(* IEC 61131-3 sources: volt/packages/volt-lsp-iec/test-corpus/bakon-nano/Device/Plc Logic/Application/Library Manager/StringUtils, 84 files *)

(* ---- CHARBUFFERPTR.dut ---- *)
TYPE CHARBUFFERPTR : POINTER TO BYTE;
END_TYPE

(* ---- DATETIMEPLACEHOLDEROCCURRENCE.dut ---- *)
TYPE DATETIMEPLACEHOLDEROCCURRENCE :
STRUCT
	M_EPLACEHOLDER : EDateTimePlaceholder;
	M_IOFFSET : INT;
	M_ILENGTH : INT;
END_STRUCT
END_TYPE

(* ---- EDATETIMEPLACEHOLDER.dut ---- *)
TYPE EDATETIMEPLACEHOLDER :
(
	PLH_IS_VALID := 0,
	DFMT_5_DIGIT_DAY := 40,
	DFMT_4_DIGIT_DAY := 41,
	DFMT_3_DIGIT_DAY := 42,
	DFMT_2_DIGIT_DAY := 43,
	DFMT_1_DIGIT_DAY := 44,
	DFMT_3_DIGIT_DAYOFYEAR := 45,
	DFMT_4_DIGIT_MONTH := 46,
	DFMT_3_DIGIT_MONTH := 47,
	DFMT_2_DIGIT_MONTH := 48,
	DFMT_1_DIGIT_MONTH := 49,
	DFMT_4_DIGIT_YEAR := 50,
	DFMT_2_DIGIT_YEAR := 51,
	DFMT_1_DIGIT_YEAR := 52,
	TFMT_2_DIGIT_HOUR_24_HOUR_CLOCK := 60,
	TFMT_1_DIGIT_HOUR_24_HOUR_CLOCK := 61,
	TFMT_2_DIGIT_HOUR_12_HOUR_CLOCK := 62,
	TFMT_1_DIGIT_HOUR_12_HOUR_CLOCK := 63,
	TFMT_3_DIGIT_MILLISECOND := 64,
	TFMT_3_DIGIT_MICROSECOND := 65,
	TFMT_3_DIGIT_NANOSECOND := 66,
	TFMT_2_DIGIT_MINUTE := 67,
	TFMT_1_DIGIT_MINUTE := 68,
	TFMT_2_DIGIT_SECOND := 69,
	TFMT_1_DIGIT_SECOND := 70,
	TFMT_AM_PM_DESIGNATOR := 71,
	TFMT_1_DIGIT_AM_PM_DESIGNATOR := 72,
	TFMT_1_DIGIT_ZONE_DESIGNATOR := 73,
	PLH_NOT_USED := 255
);
END_TYPE

(* ---- EPLACEHOLDERANALYZATIONSTATE.dut ---- *)
TYPE EPLACEHOLDERANALYZATIONSTATE :
(
	NOTAVAILABLE := 16#0,
	TOOMANYPLACEHOLDERS := 16#1,
	DONE := 16#10
);
END_TYPE

(* ---- PLACEHOLDERDESCRIPTION.dut ---- *)
TYPE PLACEHOLDERDESCRIPTION :
STRUCT
	M_EPLACEHOLDER : EDateTimePlaceholder;
	M_PCBSPLACEHOLDER : POINTER TO CharBufferString;
	M_XCONSIDERPLACEHOLDER : BOOL := TRUE;
	M_PRELATEDPLACEHOLDERISSUBSTRINGOF : POINTER TO PlaceholderDescription;
	M_PRELATEDPLACEHOLDERHASSUBSTRING : POINTER TO PlaceholderDescription;
END_STRUCT
END_TYPE

(* ---- CONSTANTS.gvl ---- *)
VAR_GLOBAL
	NULL : POINTER TO BYTE := 0;
END_VAR

(* ---- GVL_UTF8.gvl ---- *)
VAR_GLOBAL
	TRAILINGBYTESFORUTF8 : ARRAY [0..255] OF BYTE := [0, 0, 0, 0, 0, 0, 0, 0, 0, 0, 0, 0, 0, 0, 0, 0, 0, 0, 0, 0, 0, 0, 0, 0, 0, 0, 0, 0, 0, 0, 0, 0, 0, 0, 0, 0, 0, 0, 0, 0, 0, 0, 0, 0, 0, 0, 0, 0, 0, 0, 0, 0, 0, 0, 0, 0, 0, 0, 0, 0, 0, 0, 0, 0, 0, 0, 0, 0, 0, 0, 0, 0, 0, 0, 0, 0, 0, 0, 0, 0, 0, 0, 0, 0, 0, 0, 0, 0, 0, 0, 0, 0, 0, 0, 0, 0, 0, 0, 0, 0, 0, 0, 0, 0, 0, 0, 0, 0, 0, 0, 0, 0, 0, 0, 0, 0, 0, 0, 0, 0, 0, 0, 0, 0, 0, 0, 0, 0, 0, 0, 0, 0, 0, 0, 0, 0, 0, 0, 0, 0, 0, 0, 0, 0, 0, 0, 0, 0, 0, 0, 0, 0, 0, 0, 0, 0, 0, 0, 0, 0, 0, 0, 0, 0, 0, 0, 0, 0, 0, 0, 0, 0, 0, 0, 0, 0, 0, 0, 0, 0, 0, 0, 0, 0, 0, 0, 0, 0, 0, 0, 0, 0, 1, 1, 1, 1, 1, 1, 1, 1, 1, 1, 1, 1, 1, 1, 1, 1, 1, 1, 1, 1, 1, 1, 1, 1, 1, 1, 1, 1, 1, 1, 1, 1, 2, 2, 2, 2, 2, 2, 2, 2, 2, 2, 2, 2, 2, 2, 2, 2, 3, 3, 3, 3, 3, 3, 3, 3, 4, 4, 4, 4, 5, 5, 5, 5];
	FIRSTBYTEMARK : ARRAY [0..6] OF BYTE := [16#0, 16#0, 16#C0, 16#E0, 16#F0, 16#F8, 16#FC];
	OFFSETSFROMUTF8 : ARRAY [0..5] OF DWORD := [16#0, 16#3080, 16#E2080, 16#3C82080, 16#FA082080, 16#82082080];
	HALFSHIFT : INT := 10;
	HALFBASE : DWORD := 16#10000;
	HALFMASK : DWORD := 16#3FF;
	UNI_REPLACEMENT_CHAR : DWORD := 16#FFFD;
	UNI_MAX_BMP : DWORD := 16#FFFF;
	UNI_MAX_UTF16 : DWORD := 16#10FFFF;
	UNI_MAX_UTF32 : DWORD := 16#7FFFFFFF;
	UNI_MAX_LEGAL_UTF32 : DWORD := 16#10FFFF;
	BYTEMASK : DWORD := 16#BF;
	BYTEMARK : DWORD := 16#80;
	UNI_SUR_HIGH_START : DWORD := 16#D800;
	UNI_SUR_HIGH_END : DWORD := 16#DBFF;
	UNI_SUR_LOW_START : DWORD := 16#DC00;
	UNI_SUR_LOW_END : DWORD := 16#DFFF;
	ERR_SOURCE_EXHAUSTED : UDINT := 16#40A0;
	ERR_TARGET_EXHAUSTED : UDINT := 16#40A1;
	ERR_SOURCE_ILLEGAL : UDINT := 16#40A2;
END_VAR

(* ---- PLACEHOLDERCONSTANTS.gvl ---- *)
VAR_GLOBAL
	DFMT_FIRST_PLACEHOLDER : EDateTimePlaceholder := EDateTimePlaceholder.DFMT_5_DIGIT_DAY;
	DFMT_LAST_PLACEHOLDER : EDateTimePlaceholder := EDateTimePlaceholder.DFMT_1_DIGIT_YEAR;
	TFMT_FIRST_PLACEHOLDER : EDateTimePlaceholder := EDateTimePlaceholder.TFMT_2_DIGIT_HOUR_24_HOUR_CLOCK;
	TFMT_LAST_PLACEHOLDER : EDateTimePlaceholder := EDateTimePlaceholder.TFMT_1_DIGIT_ZONE_DESIGNATOR;
END_VAR

(* ---- STRINGUTILSVERSIONCONSTANTS.gvl ---- *)
VAR_GLOBAL
	_STRINGUTILS_VERSION_LARGEROREQUAL_3_5_3_40_ : INT := 0;
END_VAR

(* ---- ICHARBUFFERSTRING.itf ---- *)
INTERFACE ICHARBUFFERSTRING
END_INTERFACE

METHOD ASWSTRING : CharBufferPtr
END_METHOD

METHOD COPY : DINT
VAR_INPUT
	CBSSOURCE : REFERENCE TO CharBufferString;
END_VAR
END_METHOD

METHOD FROMSTRING : BOOL
VAR_INPUT
	STSTRING : STRING(255);
END_VAR
END_METHOD

METHOD INITCONVERTED : BOOL
VAR_INPUT
	PBUFFER : POINTER TO BYTE;
	UIBUFFERSIZE : UINT;
END_VAR
END_METHOD

(* ---- ILOCALIZEDDATETIMENAMES.itf ---- *)
INTERFACE ILOCALIZEDDATETIMENAMES
END_INTERFACE

METHOD GETDAYLONG : CharBufferPtr
VAR_INPUT
	UIDAYOFWEEK : UINT;
END_VAR
END_METHOD

METHOD GETDAYSHORT : CharBufferPtr
VAR_INPUT
	UIDAYOFWEEK : UINT;
END_VAR
END_METHOD

METHOD GETMONTHLONG : CharBufferPtr
VAR_INPUT
	UIMONTH : UINT;
END_VAR
END_METHOD

METHOD GETMONTHSHORT : CharBufferPtr
VAR_INPUT
	UIMONTH : UINT;
END_VAR
END_METHOD

(* ---- _PRINTF.pou ---- *)
FUNCTION _PRINTF : BOOL
VAR_INPUT
	CBPRESULT : CharBufferPtr;
	UIRESULTCAPACITY : UINT;
	STRINGTYPE : __SYSTEM.TYPE_CLASS;
	CBPFORMAT : CharBufferPtr;
	PVALUE : POINTER TO BYTE;
	TYPECLASS : __SYSTEM.TYPE_CLASS;
END_VAR
END_FUNCTION

(* ---- ANALYZEPLACEHOLDERS.pou ---- *)
FUNCTION ANALYZEPLACEHOLDERS : EPlaceholderAnalyzationState
VAR_INPUT
	RCBSMESSAGE : REFERENCE TO CharBufferString;
	PAPLACEHOLDERS : POINTER TO ARRAY [0..0] OF PlaceholderDescription;
	ICOUNTPLACEHOLDERTOCHECK : INT;
	PAPLACEHOLDEROCCURRENCE : POINTER TO ARRAY [0..0] OF DateTimePlaceholderOccurrence;
	SIMAXCOUNTPLACEHOLDERS : SINT;
END_VAR
VAR_OUTPUT
	SICOUNTPLACEHOLDERS : SINT;
END_VAR
END_FUNCTION

(* ---- ANALYZEPLACEHOLDERSDATETIME.pou ---- *)
FUNCTION ANALYZEPLACEHOLDERSDATETIME : EPlaceholderAnalyzationState
VAR_INPUT
	RCBSMESSAGE : REFERENCE TO CharBufferString;
	PAPLACEHOLDERS : POINTER TO ARRAY [0..0] OF PlaceholderDescription;
	ICOUNTPLACEHOLDERTOCHECK : INT;
	PAPLACEHOLDEROCCURRENCE : POINTER TO ARRAY [0..0] OF DateTimePlaceholderOccurrence;
	SIMAXCOUNTPLACEHOLDERS : SINT;
END_VAR
VAR_OUTPUT
	SICOUNTPLACEHOLDERS : SINT;
END_VAR
END_FUNCTION

(* ---- CHARACTERATEQUALS.pou ---- *)
FUNCTION CHARACTERATEQUALS : BOOL
VAR_INPUT
	CBSSOURCE : REFERENCE TO CharBufferString;
	IPOSITION : INT;
	STCHAR : STRING(1);
END_VAR
END_FUNCTION

(* ---- CHARTOUPPER.pou ---- *)
FUNCTION CHARTOUPPER : BYTE
VAR_INPUT
	BYCHAR : BYTE;
END_VAR
END_FUNCTION

(* ---- CONVERTUTF16TOUTF8.pou ---- *)
FUNCTION CONVERTUTF16TOUTF8 : UDINT
VAR_INPUT
	SOURCESTART : POINTER TO WORD;
	TARGETSTART : POINTER TO BYTE;
	DWTARGETBUFFERSIZE : DWORD;
	BSTRICTCONVERSION : BOOL;
END_VAR
END_FUNCTION

(* ---- CONVERTUTF8TOUTF16.pou ---- *)
FUNCTION CONVERTUTF8TOUTF16 : UDINT
VAR_INPUT
	SOURCESTART : POINTER TO BYTE;
	TARGETSTART : POINTER TO WORD;
	DWTARGETBUFFERSIZE : DWORD;
	BSTRICTCONVERSION : BOOL;
END_VAR
END_FUNCTION

(* ---- HELPISSAMEIGNORECASE.pou ---- *)
FUNCTION HELPISSAMEIGNORECASE : BOOL
VAR_INPUT
	BY1 : BYTE;
	BY2 : BYTE;
END_VAR
END_FUNCTION

(* ---- HELPSTRCMPENDA.pou ---- *)
FUNCTION HELPSTRCMPENDA : BOOL
VAR_INPUT
	PCOMPLETETEXT : CharBufferPtr;
	PSUBTEXT : CharBufferPtr;
	XIGNORECASE : BOOL;
END_VAR
END_FUNCTION

(* ---- HELPSTRCMPSTARTA.pou ---- *)
FUNCTION HELPSTRCMPSTARTA : BOOL
VAR_INPUT
	PCOMPLETETEXT : CharBufferPtr;
	PSUBTEXT : CharBufferPtr;
	XIGNORECASE : BOOL;
END_VAR
END_FUNCTION

(* ---- HELPTRIM.pou ---- *)
FUNCTION HELPTRIM : POINTER TO BYTE
VAR_INPUT
	PTEXT : CharBufferPtr;
	XTRIMLEFT : BOOL;
END_VAR
END_FUNCTION

(* ---- HELPTRIMW.pou ---- *)
FUNCTION HELPTRIMW : POINTER TO WORD
VAR_INPUT
	PTEXT : CharBufferPtr;
	XTRIMLEFT : BOOL;
END_VAR
END_FUNCTION

(* ---- ISLEGALUTF8.pou ---- *)
FUNCTION ISLEGALUTF8 : BOOL
VAR_INPUT
	SOURCE : POINTER TO BYTE;
	LENGTH : INT;
END_VAR
END_FUNCTION

(* ---- ISSPACECHARACTER.pou ---- *)
FUNCTION ISSPACECHARACTER : BOOL
VAR_INPUT
	WCHARACTER : WORD;
END_VAR
END_FUNCTION

(* ---- PRINTF.pou ---- *)
FUNCTION PRINTF
VAR_INPUT
	CBSRESULT : REFERENCE TO CharBufferString;
	CBSFORMAT : REFERENCE TO CharBufferString;
	PVALUE : POINTER TO BYTE;
	TYPECLASS : __SYSTEM.TYPE_CLASS;
END_VAR
END_FUNCTION

(* ---- STRATOW.pou ---- *)
FUNCTION STRATOW
VAR_INPUT
	PBYTARGETW : POINTER TO BYTE;
	IBUFFERSIZE : DINT;
	PBYSOURCEA : POINTER TO BYTE;
END_VAR
END_FUNCTION

(* ---- STRCASECMPA.pou ---- *)
FUNCTION STRCASECMPA : INT
VAR_INPUT
	PBYTE1 : POINTER TO BYTE;
	PBYTE2 : POINTER TO BYTE;
END_VAR
END_FUNCTION

(* ---- STRCASECMPENDA.pou ---- *)
FUNCTION STRCASECMPENDA : INT
VAR_INPUT
	PSTRING : CharBufferPtr;
	PSUFFIX : CharBufferPtr;
END_VAR
END_FUNCTION

(* ---- STRCASECMPSTARTA.pou ---- *)
FUNCTION STRCASECMPSTARTA : INT
VAR_INPUT
	PSTRING : CharBufferPtr;
	PPREFIX : CharBufferPtr;
END_VAR
END_FUNCTION

(* ---- STRCASECMPW.pou ---- *)
FUNCTION STRCASECMPW : INT
VAR_INPUT
	PWD1 : POINTER TO WORD;
	PWD2 : POINTER TO WORD;
END_VAR
END_FUNCTION

(* ---- STRCASEFINDA.pou ---- *)
FUNCTION STRCASEFINDA : INT
VAR_INPUT
	PST1 : POINTER TO STRING(255);
	PST2 : POINTER TO STRING(255);
	UISEARCHSTART : UINT;
END_VAR
END_FUNCTION

(* ---- STRCASEFINDW.pou ---- *)
FUNCTION STRCASEFINDW : INT
VAR_INPUT
	PST1 : POINTER TO WSTRING(255);
	PST2 : POINTER TO WSTRING(255);
	UISEARCHSTART : UINT;
END_VAR
END_FUNCTION

(* ---- STRCMP.pou ---- *)
FUNCTION STRCMP : DINT
VAR_INPUT
	CBSSTRING1 : REFERENCE TO CharBufferString;
	CBSSTRING2 : REFERENCE TO CharBufferString;
END_VAR
END_FUNCTION

(* ---- STRCMPA.pou ---- *)
FUNCTION STRCMPA : INT
VAR_INPUT
	PBY1 : POINTER TO BYTE;
	PBY2 : POINTER TO BYTE;
END_VAR
END_FUNCTION

(* ---- STRCMPENDA.pou ---- *)
FUNCTION STRCMPENDA : INT
VAR_INPUT
	PSTRING : CharBufferPtr;
	PSUFFIX : CharBufferPtr;
END_VAR
END_FUNCTION

(* ---- STRCMPSTARTA.pou ---- *)
FUNCTION STRCMPSTARTA : INT
VAR_INPUT
	PSTRING : CharBufferPtr;
	PPREFIX : CharBufferPtr;
END_VAR
END_FUNCTION

(* ---- STRCMPW.pou ---- *)
FUNCTION STRCMPW : INT
VAR_INPUT
	PWD1 : POINTER TO WORD;
	PWD2 : POINTER TO WORD;
END_VAR
END_FUNCTION

(* ---- STRCONCATA.pou ---- *)
FUNCTION STRCONCATA : BOOL
VAR_INPUT
	PSTFROM : CharBufferPtr;
	PSTTO : CharBufferPtr;
	IBUFFERSIZE : INT;
END_VAR
END_FUNCTION

(* ---- STRCONCATW.pou ---- *)
FUNCTION STRCONCATW : BOOL
VAR_INPUT
	PSTFROM : CharBufferPtr;
	PSTTO : CharBufferPtr;
	IBUFFERSIZE : INT;
END_VAR
END_FUNCTION

(* ---- STRCPY.pou ---- *)
FUNCTION STRCPY : DINT
VAR_INPUT
	CBSTARGET : REFERENCE TO CharBufferString;
	CBSSOURCE : REFERENCE TO CharBufferString;
END_VAR
END_FUNCTION

(* ---- STRCPYA.pou ---- *)
FUNCTION STRCPYA : DINT
VAR_INPUT
	PBUFFER : CharBufferPtr;
	IBUFFERSIZE : DINT;
	PSTR : CharBufferPtr;
END_VAR
END_FUNCTION

(* ---- STRCPYFROM.pou ---- *)
FUNCTION STRCPYFROM : DINT
VAR_INPUT
	RCBSTARGET : REFERENCE TO CharBufferString;
	RCBSSOURCE : REFERENCE TO CharBufferString;
	DISOURCEOFFSET : DINT;
	DITARGETOFFSET : DINT;
	DICOUNTCHARACTERS : DINT;
END_VAR
END_FUNCTION

(* ---- STRCPYW.pou ---- *)
FUNCTION STRCPYW : DINT
VAR_INPUT
	PBUFFER : CharBufferPtr;
	IBUFFERSIZE : DINT;
	PSTR : CharBufferPtr;
END_VAR
END_FUNCTION

(* ---- STRDELETE.pou ---- *)
FUNCTION STRDELETE
VAR_INPUT
	CBSSOURCE : REFERENCE TO CharBufferString;
	ILENGTH : INT;
	IPOSITION : INT;
END_VAR
END_FUNCTION

(* ---- STRDELETEA.pou ---- *)
FUNCTION STRDELETEA
VAR_INPUT
	PBY : POINTER TO BYTE;
	ILENGTH : INT;
	IPOSITION : INT;
END_VAR
END_FUNCTION

(* ---- STRDELETEW.pou ---- *)
FUNCTION STRDELETEW
VAR_INPUT
	PWD : POINTER TO WORD;
	ILENGTH : INT;
	IPOSITION : INT;
END_VAR
END_FUNCTION

(* ---- STRFIND.pou ---- *)
FUNCTION STRFIND : INT
VAR_INPUT
	CBSSOURCE : REFERENCE TO CharBufferString;
	CBSTOSEARCHFOR : REFERENCE TO CharBufferString;
END_VAR
END_FUNCTION

(* ---- STRFINDA.pou ---- *)
FUNCTION STRFINDA : INT
VAR_INPUT
	PST1 : POINTER TO STRING(255);
	PST2 : POINTER TO STRING(255);
	UISEARCHSTART : UINT;
END_VAR
END_FUNCTION

(* ---- STRFINDFROM.pou ---- *)
FUNCTION STRFINDFROM : INT
VAR_INPUT
	CBSSOURCE : REFERENCE TO CharBufferString;
	CBSTOSEARCHFOR : REFERENCE TO CharBufferString;
	ISEARCHSTART : UINT;
END_VAR
END_FUNCTION

(* ---- STRFINDW.pou ---- *)
FUNCTION STRFINDW : INT
VAR_INPUT
	PST1 : POINTER TO WSTRING(255);
	PST2 : POINTER TO WSTRING(255);
	UISEARCHSTART : UINT;
END_VAR
END_FUNCTION

(* ---- STRINGTOCHARBUFFERPTR.pou ---- *)
FUNCTION STRINGTOCHARBUFFERPTR : BOOL
VAR_INPUT
	STSTRING : STRING(255);
	CBSRESULT : REFERENCE TO CharBufferString;
END_VAR
END_FUNCTION

(* ---- STRINSERT.pou ---- *)
FUNCTION STRINSERT
VAR_INPUT
	CBSINPUT : REFERENCE TO CharBufferString;
	CBSINSERT : REFERENCE TO CharBufferString;
	IPOSITION : INT;
END_VAR
END_FUNCTION

(* ---- STRISNULLOREMPTYA.pou ---- *)
FUNCTION STRISNULLOREMPTYA : BOOL
VAR_INPUT
	PSTDATA : CharBufferPtr;
END_VAR
END_FUNCTION

(* ---- STRISNULLOREMPTYW.pou ---- *)
FUNCTION STRISNULLOREMPTYW : BOOL
VAR_INPUT
	PSTDATA : CharBufferPtr;
END_VAR
END_FUNCTION

(* ---- STRLEN.pou ---- *)
FUNCTION STRLEN : DINT
VAR_INPUT
	CBSSOURCE : REFERENCE TO CharBufferString;
END_VAR
END_FUNCTION

(* ---- STRLENA.pou ---- *)
FUNCTION STRLENA : DINT
VAR_INPUT
	PSTDATA : CharBufferPtr;
END_VAR
END_FUNCTION

(* ---- STRLENW.pou ---- *)
FUNCTION STRLENW : DINT
VAR_INPUT
	PSTDATA : CharBufferPtr;
END_VAR
END_FUNCTION

(* ---- STRMID.pou ---- *)
FUNCTION STRMID
VAR_INPUT
	CBSSOURCE : REFERENCE TO CharBufferString;
	ILENGTH : INT;
	IPOSITION : INT;
	CBSRESULT : REFERENCE TO CharBufferString;
END_VAR
END_FUNCTION

(* ---- STRMIDA.pou ---- *)
FUNCTION STRMIDA
VAR_INPUT
	PST : POINTER TO BYTE;
	UIINPUTBUFFERSIZE : UINT;
	ILENGTH : INT;
	IPOSITION : INT;
	PSTRESULT : POINTER TO BYTE;
	UIRESULTBUFFERSIZE : UINT;
END_VAR
END_FUNCTION

(* ---- STRMIDW.pou ---- *)
FUNCTION STRMIDW
VAR_INPUT
	PWST : POINTER TO WORD;
	UIINPUTBUFFERSIZE : UINT;
	ILENGTH : INT;
	IPOSITION : INT;
	PWSTRESULT : POINTER TO WORD;
	UIRESULTBUFFERSIZE : UINT;
END_VAR
END_FUNCTION

(* ---- STRPADLEFTA.pou ---- *)
FUNCTION STRPADLEFTA : BOOL
VAR_INPUT
	BYPADCHAR : BYTE;
	PSTFROM : CharBufferPtr;
	PSTTO : CharBufferPtr;
	DIBUFFERSIZE : DINT;
END_VAR
END_FUNCTION

(* ---- STRPADLEFTW.pou ---- *)
FUNCTION STRPADLEFTW : BOOL
VAR_INPUT
	WPADCHAR : WORD;
	PSTFROM : CharBufferPtr;
	PSTTO : CharBufferPtr;
	DIBUFFERSIZE : DINT;
END_VAR
END_FUNCTION

(* ---- STRPADRIGHTA.pou ---- *)
FUNCTION STRPADRIGHTA : BOOL
VAR_INPUT
	BYPADCHAR : BYTE;
	PSTFROM : CharBufferPtr;
	PSTTO : CharBufferPtr;
	DIBUFFERSIZE : DINT;
END_VAR
END_FUNCTION

(* ---- STRPADRIGHTW.pou ---- *)
FUNCTION STRPADRIGHTW : BOOL
VAR_INPUT
	WPADCHAR : WORD;
	PSTFROM : CharBufferPtr;
	PSTTO : CharBufferPtr;
	DIBUFFERSIZE : DINT;
END_VAR
END_FUNCTION

(* ---- STRREPLACE.pou ---- *)
FUNCTION STRREPLACE
VAR_INPUT
	CBSINPUT : REFERENCE TO CharBufferString;
	CBSREPLACEWITH : REFERENCE TO CharBufferString;
	ILENGTHTOREPLACE : INT;
	IPOSITION : INT;
END_VAR
END_FUNCTION

(* ---- STRREPLACEA.pou ---- *)
FUNCTION STRREPLACEA
VAR_INPUT
	PSTINPUT : POINTER TO STRING(255);
	UIINPUTBUFFERSIZE : UINT;
	PSTREPLACEWITH : POINTER TO STRING(255);
	ILENGTHINPUT : INT;
	ILENGTHTOREPLACE : INT;
	ILENGTHTOREPLACEWITH : INT;
	IPOSITION : INT;
END_VAR
END_FUNCTION

(* ---- STRREPLACEW.pou ---- *)
FUNCTION STRREPLACEW
VAR_INPUT
	PSTINPUT : POINTER TO WSTRING(255);
	UIINPUTBUFFERSIZE : UINT;
	PSTREPLACEWITH : POINTER TO WSTRING(255);
	ILENGTHINPUT : INT;
	ILENGTHTOREPLACE : INT;
	ILENGTHTOREPLACEWITH : INT;
	IPOSITION : INT;
END_VAR
END_FUNCTION

(* ---- STRTOLOWERA.pou ---- *)
FUNCTION STRTOLOWERA
VAR_INPUT
	PSTRING : CharBufferPtr;
END_VAR
END_FUNCTION

(* ---- STRTOUPPERA.pou ---- *)
FUNCTION STRTOUPPERA
VAR_INPUT
	PSTRING : CharBufferPtr;
END_VAR
END_FUNCTION

(* ---- STRTRIMA.pou ---- *)
FUNCTION STRTRIMA
VAR_INPUT
	PSTRING : POINTER TO BYTE;
END_VAR
END_FUNCTION

(* ---- STRTRIMENDA.pou ---- *)
FUNCTION STRTRIMENDA
VAR_INPUT
	PSTRING : POINTER TO BYTE;
END_VAR
END_FUNCTION

(* ---- STRTRIMENDW.pou ---- *)
FUNCTION STRTRIMENDW
VAR_INPUT
	PSTRING : CharBufferPtr;
END_VAR
END_FUNCTION

(* ---- STRTRIMSTARTA.pou ---- *)
FUNCTION STRTRIMSTARTA
VAR_INPUT
	PSTRING : POINTER TO BYTE;
END_VAR
END_FUNCTION

(* ---- STRTRIMSTARTW.pou ---- *)
FUNCTION STRTRIMSTARTW
VAR_INPUT
	PSTRING : CharBufferPtr;
END_VAR
END_FUNCTION

(* ---- STRTRIMW.pou ---- *)
FUNCTION STRTRIMW : BOOL
VAR_INPUT
	PSTRING : CharBufferPtr;
END_VAR
END_FUNCTION

(* ---- STUSPRINTF.pou ---- *)
FUNCTION STUSPRINTF : INT
VAR_INPUT
	PSTFORMAT : POINTER TO STRING;
	PVARADR : POINTER TO DWORD;
	UDIVARTYPE : __SYSTEM.TYPE_CLASS;
	PBUFFER : POINTER TO BYTE;
	DWBUFFERSIZE : UDINT;
END_VAR
END_FUNCTION

(* ---- STUSPRINTFW.pou ---- *)
FUNCTION STUSPRINTFW : INT
VAR_INPUT
	WSTFORMAT : POINTER TO WSTRING;
	PVARADR : POINTER TO DWORD;
	UDIVARTYPE : __SYSTEM.TYPE_CLASS;
	PBUFFER : POINTER TO BYTE;
	DWBUFFERSIZE : UDINT;
END_VAR
END_FUNCTION

(* ---- WCHARTOUPPER.pou ---- *)
FUNCTION WCHARTOUPPER : WORD
VAR_INPUT
	WDCHAR : WORD;
END_VAR
END_FUNCTION

(* ---- ABSTRACTFORMATTER.pou ---- *)
FUNCTION_BLOCK ABSTRACTFORMATTER
VAR
	M_APLACEHOLDEROCCURRENCE : ARRAY [0..(COUNT_PLACEHOLDERS_IN_FORMAT_STRING - 1)] OF DateTimePlaceholderOccurrence;
	M_SICOUNTPLACEHOLDERS : SINT := -1;
	M_EPLACEHOLDERANALYZATIONSTATE : EPlaceholderAnalyzationState;
	M_SFORMATSTRING : STRING(50);
	M_IFORMATSTRINGLENGTH : INT;
	COUNT_PLACEHOLDERS_IN_FORMAT_STRING : INT := 10;
	COUNT_PLACEHOLDERS_IN_DATETIMEFORMAT_STRING : INT := 20;
	MAX_FORMAT_STRING_LENGTH : SINT := 50;
END_VAR
END_FUNCTION_BLOCK

(* ---- CHARBUFFERSTRING.pou ---- *)
FUNCTION_BLOCK CHARBUFFERSTRING
VAR_INPUT
	M_UIBUFFERSIZE : UINT;
	M_CBPBUFFER : CharBufferPtr;
	M_TYPE : __SYSTEM.TYPE_CLASS;
	M_ASSTRING : POINTER TO STRING(255);
	M_ASWSTRING : POINTER TO WSTRING(255);
	M_BALLOCATED : BOOL;
END_VAR
VAR
	CAPACITY : UINT;
	CHARACTERS : CharBufferPtr;
	LENGTH : DINT;
	STRINGTYPE : __SYSTEM.TYPE_CLASS;
END_VAR
END_FUNCTION_BLOCK

METHOD ASWSTRING : CharBufferPtr
END_METHOD

METHOD CHARAT : BYTE
VAR_INPUT
	IPOSITION : INT;
END_VAR
END_METHOD

METHOD CHARATEQUALS : BOOL
VAR_INPUT
	IPOSITION : INT;
	STCHAR : STRING(1);
END_VAR
END_METHOD

METHOD COPY : DINT
VAR_INPUT
	CBSSOURCE : REFERENCE TO CharBufferString;
END_VAR
END_METHOD

METHOD COPYFROM
VAR_INPUT
	RCBSSOURCE : REFERENCE TO CharBufferString;
	DISOURCEOFFSET : DINT;
	DITARGETOFFSET : DINT;
	DICOUNTCHARACTERS : DINT;
END_VAR
END_METHOD

METHOD COPYFROM2 : DINT
VAR_INPUT
	RSSOURCE : REFERENCE TO STRING(255);
	DITARGETOFFSET : DINT;
END_VAR
END_METHOD

METHOD DELETE : DINT
VAR_INPUT
	ILENGTH : INT;
	IPOSITION : INT;
END_VAR
END_METHOD

METHOD FB_EXIT : BOOL
VAR_INPUT
	BINCOPYCODE : BOOL;
END_VAR
END_METHOD

METHOD FB_INIT : BOOL
VAR_INPUT
	BINITRETAINS : BOOL;
	BINCOPYCODE : BOOL;
	UIBUFFERSIZE : UINT;
	STRINGTYPE : __SYSTEM.TYPE_CLASS;
END_VAR
END_METHOD

METHOD FIND : INT
VAR_INPUT
	CBSTOSEARCHFOR : REFERENCE TO CharBufferString;
END_VAR
END_METHOD

METHOD FINDFROM : INT
VAR_INPUT
	CBSTOSEARCHFOR : REFERENCE TO CharBufferString;
	ISEARCHSTART : UINT;
END_VAR
END_METHOD

METHOD FROMSTRING : BOOL
VAR_INPUT
	STSTRING : STRING(255);
END_VAR
END_METHOD

METHOD INIT : BOOL
VAR_INPUT
	PBUFFER : POINTER TO BYTE;
	UIBUFFERSIZE : UINT;
	STRINGTYPE : __SYSTEM.TYPE_CLASS;
END_VAR
END_METHOD

METHOD INITCONVERTED : BOOL
VAR_INPUT
	PBUFFER : POINTER TO BYTE;
	UIBUFFERSIZE : UINT;
END_VAR
END_METHOD

METHOD INITIALIZE : BOOL
VAR_INPUT
	CBPSOURCE : CharBufferPtr;
	STRINGTYPE : __SYSTEM.TYPE_CLASS;
END_VAR
END_METHOD

METHOD INSERT
VAR_INPUT
	CBSINSERT : REFERENCE TO CharBufferString;
	IPOSITION : INT;
END_VAR
END_METHOD

METHOD MID
VAR_INPUT
	ILENGTH : INT;
	IPOSITION : INT;
	CBSRESULT : REFERENCE TO CharBufferString;
END_VAR
END_METHOD

METHOD PLACEHOLDEREQUALS : BOOL
VAR_INPUT
	STVALUE : STRING;
	WSTVALUE : WSTRING;
END_VAR
END_METHOD

METHOD REPLACE
VAR_INPUT
	CBSREPLACEWITH : REFERENCE TO CharBufferString;
	ILENGTHTOREPLACE : INT;
	IPOSITION : INT;
END_VAR
END_METHOD

(* ---- DATEFORMATTER.pou ---- *)
FUNCTION_BLOCK DATEFORMATTER EXTENDS AbstractFormatter
VAR
	M_CBSPLACEHOLDER2DIGITDAY : CharBufferString;
	M_CBSPLACEHOLDER1DIGITDAY : CharBufferString;
	M_CBSPLACEHOLDER2DIGITMONTH : CharBufferString;
	M_CBSPLACEHOLDER1DIGITMONTH : CharBufferString;
	M_CBSPLACEHOLDER4DIGITYEAR : CharBufferString;
	M_CBSPLACEHOLDER2DIGITYEAR : CharBufferString;
	M_CBSPLACEHOLDER1DIGITYEAR : CharBufferString;
END_VAR
END_FUNCTION_BLOCK

METHOD FB_EXIT : BOOL
VAR_INPUT
	BINCOPYCODE : BOOL;
END_VAR
END_METHOD

METHOD FB_INIT : BOOL
VAR_INPUT
	BINITRETAINS : BOOL;
	BINCOPYCODE : BOOL;
END_VAR
END_METHOD

METHOD FORMAT : STRING
VAR_INPUT
	PDATE : SYSTIMEDATE;
END_VAR
END_METHOD

METHOD SETFORMATSTRING
VAR_INPUT
	SFORMATSTRING : STRING(MAX_FORMAT_STRING_LENGTH);
END_VAR
END_METHOD

(* ---- DATETIMEFORMATTER.pou ---- *)
FUNCTION_BLOCK DATETIMEFORMATTER EXTENDS AbstractFormatter
VAR
	M_APLACEHOLDEROCCURRENCEDATETIME : ARRAY [0..(COUNT_PLACEHOLDERS_IN_DATETIMEFORMAT_STRING - 1)] OF DateTimePlaceholderOccurrence;
	M_CBSPLACEHOLDER5DIGITDAY : CharBufferString;
	M_CBSPLACEHOLDER4DIGITDAY : CharBufferString;
	M_CBSPLACEHOLDER3DIGITDAY : CharBufferString;
	M_CBSPLACEHOLDER2DIGITDAY : CharBufferString;
	M_CBSPLACEHOLDER1DIGITDAY : CharBufferString;
	M_CBSPLACEHOLDER3DIGITDAYOFYEAR : CharBufferString;
	M_CBSPLACEHOLDER4DIGITMONTH : CharBufferString;
	M_CBSPLACEHOLDER3DIGITMONTH : CharBufferString;
	M_CBSPLACEHOLDER2DIGITMONTH : CharBufferString;
	M_CBSPLACEHOLDER1DIGITMONTH : CharBufferString;
	M_CBSPLACEHOLDER4DIGITYEAR : CharBufferString;
	M_CBSPLACEHOLDER2DIGITYEAR : CharBufferString;
	M_CBSPLACEHOLDER1DIGITYEAR : CharBufferString;
	M_CBSPLACEHOLDER2DIGITHOUR24HOURCLOCK : CharBufferString;
	M_CBSPLACEHOLDER1DIGITHOUR24HOURCLOCK : CharBufferString;
	M_CBSPLACEHOLDER2DIGITHOUR12HOURCLOCK : CharBufferString;
	M_CBSPLACEHOLDER1DIGITHOUR12HOURCLOCK : CharBufferString;
	M_CBSPLACEHOLDER2DIGITMINUTE : CharBufferString;
	M_CBSPLACEHOLDER1DIGITMINUTE : CharBufferString;
	M_CBSPLACEHOLDER2DIGITSECOND : CharBufferString;
	M_CBSPLACEHOLDER1DIGITSECOND : CharBufferString;
	M_CBSPLACEHOLDER3DIGITMILLISECOND : CharBufferString;
	M_CBSPLACEHOLDER3DIGITMICROSECOND : CharBufferString;
	M_CBSPLACEHOLDER3DIGITNANOSECOND : CharBufferString;
	M_CBSPLACEHOLDER2DIGITAMPMDESIGNATOR : CharBufferString;
	M_CBSPLACEHOLDER1DIGITAMPMDESIGNATOR : CharBufferString;
	M_CBSPLACEHOLDER1DIGITZONEDESIGNATOR : CharBufferString;
	M_OPTLOCALIZER : ILocalizedDateTimeNames;
	M_IUTCOFFSET : INT;
END_VAR
END_FUNCTION_BLOCK

METHOD FB_EXIT : BOOL
VAR_INPUT
	BINCOPYCODE : BOOL;
END_VAR
END_METHOD

METHOD FB_INIT : BOOL
VAR_INPUT
	BINITRETAINS : BOOL;
	BINCOPYCODE : BOOL;
END_VAR
END_METHOD

METHOD FORMAT : WSTRING
VAR_INPUT
	PDATE : SYSTIMEDATE;
	UIMICROSECONDS : UINT;
	UINANOSECONDS : UINT;
	DATATYPE : __SYSTEM.TYPE_CLASS := __SYSTEM.TYPE_CLASS.TYPE_NONE;
END_VAR
END_METHOD

METHOD FORMATSINGLEDIGIT : WSTRING
VAR_INPUT
	PDATE : SYSTIMEDATE;
	UIMICROSECONDS : UINT;
	UINANOSECONDS : UINT;
	DATATYPE : __SYSTEM.TYPE_CLASS := __SYSTEM.TYPE_CLASS.TYPE_NONE;
	SIINDEXOFSINGLEDIGITTORETURN : SINT;
END_VAR
VAR_OUTPUT
	ICOPYSINGLETARGETOFFSET : INT;
END_VAR
END_METHOD

METHOD FORMATWITHUTCOFFSET : WSTRING
VAR_INPUT
	PDATE : SYSTIMEDATE;
	UIMICROSECONDS : UINT;
	UINANOSECONDS : UINT;
	DATATYPE : __SYSTEM.TYPE_CLASS := __SYSTEM.TYPE_CLASS.TYPE_NONE;
	IUTCOFFSET : INT;
END_VAR
END_METHOD

METHOD SETFORMATSTRING
VAR_INPUT
	SFORMATSTRING : STRING(MAX_FORMAT_STRING_LENGTH);
END_VAR
END_METHOD

METHOD SETLOCALIZER
VAR_INPUT
	LOCALIZER : ILocalizedDateTimeNames;
END_VAR
END_METHOD

METHOD GETDAY : WSTRING
VAR_INPUT
	UIDAYOFWEEK : UINT;
	DAYFORMAT : EDateTimePlaceholder;
END_VAR
VAR_IN_OUT
	DILENGTH : DINT;
END_VAR
END_METHOD

METHOD GETMONTH : WSTRING
VAR_INPUT
	UIMONTH : UINT;
	MONTHFORMAT : EDateTimePlaceholder;
END_VAR
VAR_IN_OUT
	DILENGTH : DINT;
END_VAR
END_METHOD

(* ---- TIMEFORMATTER.pou ---- *)
FUNCTION_BLOCK TIMEFORMATTER EXTENDS AbstractFormatter
VAR
	M_CBSPLACEHOLDER2DIGITHOUR24HOURCLOCK : CharBufferString;
	M_CBSPLACEHOLDER1DIGITHOUR24HOURCLOCK : CharBufferString;
	M_CBSPLACEHOLDER2DIGITHOUR12HOURCLOCK : CharBufferString;
	M_CBSPLACEHOLDER1DIGITHOUR12HOURCLOCK : CharBufferString;
	M_CBSPLACEHOLDER2DIGITMINUTE : CharBufferString;
	M_CBSPLACEHOLDER1DIGITMINUTE : CharBufferString;
	M_CBSPLACEHOLDER2DIGITSECOND : CharBufferString;
	M_CBSPLACEHOLDER1DIGITSECOND : CharBufferString;
	M_CBSPLACEHOLDER3DIGITMILLISECOND : CharBufferString;
	M_CBSPLACEHOLDER3DIGITMICROSECOND : CharBufferString;
	M_CBSPLACEHOLDERAMPMDESIGNATOR : CharBufferString;
	M_CBSPLACEHOLDER1DIGITZONEDESIGNATOR : CharBufferString;
END_VAR
END_FUNCTION_BLOCK

METHOD FB_EXIT : BOOL
VAR_INPUT
	BINCOPYCODE : BOOL;
END_VAR
END_METHOD

METHOD FB_INIT : BOOL
VAR_INPUT
	BINITRETAINS : BOOL;
	BINCOPYCODE : BOOL;
END_VAR
END_METHOD

METHOD FORMAT : STRING
VAR_INPUT
	PDATE : SYSTIMEDATE;
	UIMIRCOSECONDS : UINT;
END_VAR
END_METHOD

METHOD FORMATWITHUTCOFFSET : STRING
VAR_INPUT
	PDATE : SYSTIMEDATE;
	UIMIRCOSECONDS : UINT;
	IUTCOFFSET : INT;
END_VAR
END_METHOD

METHOD SETFORMATSTRING
VAR_INPUT
	SFORMATSTRING : STRING(MAX_FORMAT_STRING_LENGTH);
END_VAR
END_METHOD
